// TIA Portal V21 export
FUNCTION_BLOCK "FB_LadBoxes"   // FB7, LAD
TITLE = LAD boxes, call and jump
{ S7_Optimized_Access := 'TRUE' }
// stored: MemoryReserve 100, SetENOAutomatically false
   VAR_INPUT
      Start : Bool;   // Start command
      InValue : Int;   // Input value
      Limit : Int := 100;   // Limit for the comparisons
   END_VAR
   VAR_OUTPUT
      Delayed : Bool;   // Start delayed by three seconds
      Copy : Int;   // Copy of the input value
      Sum : Int;   // Input value plus limit
      IsEqual : Bool;   // Input value equal to the limit
      IsGreater : Bool;   // Input value greater than the limit
      IsLessEqual : Bool;   // Input value less than or equal to the limit
      Average : Real;   // Average from FB_SclSections
      SectionsOk : Bool;   // ENO of the FB_SclSections call
      Skipped : Bool;   // Set only when the jump is not taken
      AfterJump : Bool;   // Network after the jump label
   END_VAR
   VAR
      Delay { S7_SetPoint := 'True'} : TON_TIME;   // On-delay timer
      DelayElapsed : Time;   // Elapsed time of the on-delay timer
      Sections { S7_SetPoint := 'True'} : "FB_SclSections";   // Multi-instance of FB_SclSections
      Values : Array[0..9] of Real;   // Values for FB_SclSections
      SectionsBusy : Bool;   // Busy output of FB_SclSections
      SectionsSteps : Int;   // Step count of FB_SclSections
      Setpoint : Real := 50.0;   // Setpoint for FB_SclSections
   END_VAR
   VAR_TEMP   // added for the SCL form of the ladder/FBD networks
      _w1 : Bool;
   END_VAR
BEGIN

REGION Network 1: On-delay timer as multi-instance
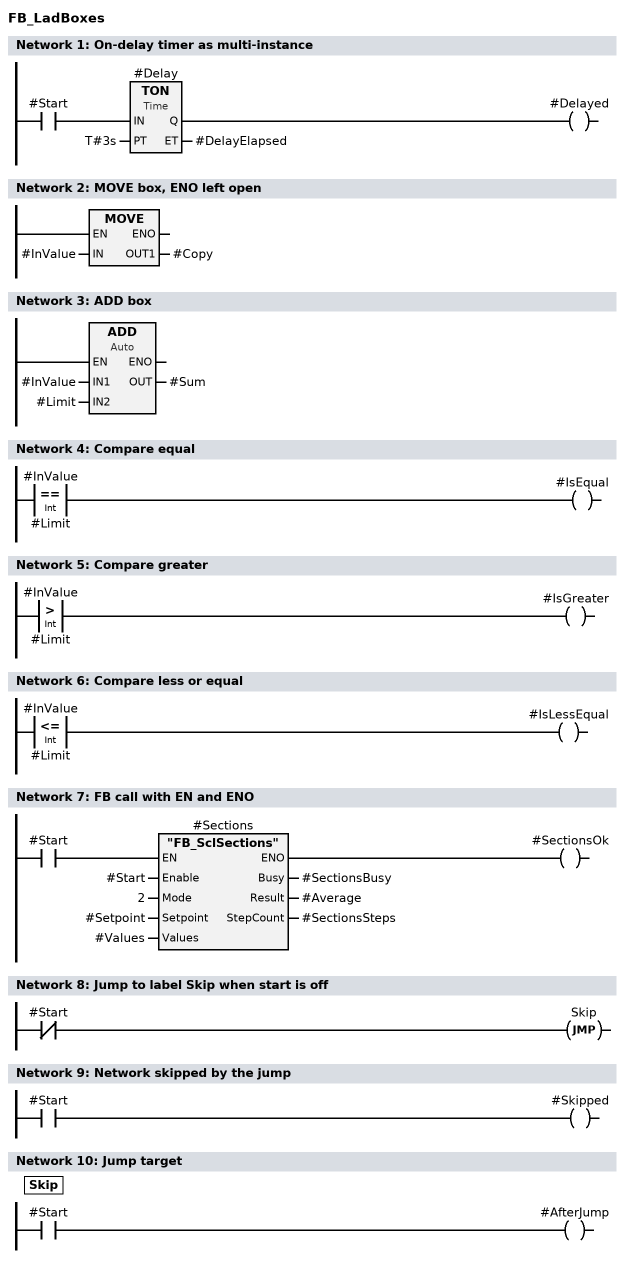
   RUNG wire#powerrail
      Contact( #Start )
      { S7_Templates := "time_type := Time" } #Delay.TON(pt := T#3s, et => #DelayElapsed)
      Coil( #Delayed )
   END_RUNG
   // the same network as SCL:
   #Delay(IN := #Start, PT := T#3s, ET => #DelayElapsed);   // TON
   #Delayed := #Delay.Q;
END_REGION

REGION Network 2: MOVE box, ENO left open
   RUNG wire#powerrail
      Move(in := #InValue, out1 => #Copy)
   END_RUNG
   // the same network as SCL:
   #Copy := #InValue;
END_REGION

REGION Network 3: ADD box
   RUNG wire#powerrail
      Add(in1 := #InValue, in2 := #Limit, out => #Sum)
   END_RUNG
   // the same network as SCL:
   #Sum := #InValue + #Limit;
END_REGION

REGION Network 4: Compare equal
   RUNG wire#powerrail
      { S7_Templates := "SrcType := Int" } EQ_Contact(in1 := #InValue, in2 := #Limit)
      Coil( #IsEqual )
   END_RUNG
   // the same network as SCL:
   #IsEqual := #InValue = #Limit;
END_REGION

REGION Network 5: Compare greater
   RUNG wire#powerrail
      { S7_Templates := "SrcType := Int" } GT_Contact(in1 := #InValue, in2 := #Limit)
      Coil( #IsGreater )
   END_RUNG
   // the same network as SCL:
   #IsGreater := #InValue > #Limit;
END_REGION

REGION Network 6: Compare less or equal
   RUNG wire#powerrail
      { S7_Templates := "SrcType := Int" } LE_Contact(in1 := #InValue, in2 := #Limit)
      Coil( #IsLessEqual )
   END_RUNG
   // the same network as SCL:
   #IsLessEqual := #InValue <= #Limit;
END_REGION

REGION Network 7: FB call with EN and ENO
   RUNG wire#powerrail
      Contact( #Start )
      #Sections(Enable := #Start, Mode := 2, Setpoint := #Setpoint, Busy => #SectionsBusy, Result => #Average, StepCount => #SectionsSteps, Values := #Values)
      Coil( #SectionsOk )
   END_RUNG
   // the same network as SCL:
   #Sections(EN := #Start,   // "FB_SclSections"
             Enable := #Start,
             Mode := 2,
             Setpoint := #Setpoint,
             Values := #Values,
             Busy => #SectionsBusy,
             Result => #Average,
             StepCount => #SectionsSteps,
             ENO => #_w1);
   #SectionsOk := #_w1;
END_REGION

REGION Network 8: Jump to label Skip when start is off
   RUNG wire#powerrail
      I_Contact( #Start )
      JumpCoil( Skip )
   END_RUNG
   // the same network as SCL:
   IF NOT #Start THEN GOTO Skip; END_IF;
END_REGION

REGION Network 9: Network skipped by the jump
   RUNG wire#powerrail
      Contact( #Start )
      Coil( #Skipped )
   END_RUNG
   // the same network as SCL:
   #Skipped := #Start;
END_REGION

REGION Network 10: Jump target
   Label( Skip )
   RUNG wire#powerrail
      Contact( #Start )
      Coil( #AfterJump )
   END_RUNG
   // the same network as SCL:
   Skip:
   #AfterJump := #Start;
END_REGION
END_FUNCTION_BLOCK
